TYPE "NameItem"
STRUCT
  Value : INT;
END_STRUCT;
END_TYPE
